// TIA Portal V20 export
// export: Created 2026-10-20T18:56:01.9058217Z, ExportSetting None, DisplayName Totally Integrated Automation Portal, DisplayVersion V20 Update 6, DisplayName TIA Portal Openness, DisplayVersion V20 Update 6, DisplayName TIA Portal Version Control Interface, DisplayVersion V20 Update 6, DisplayName SINAMICS Startdrive Advanced, DisplayVersion V20 SP1, DisplayName SINAMICS Startdrive G130, G150, S120, S150, SINAMICS MV, G220, S200, S210, DisplayVersion V20 SP1, DisplayName SINAMICS Startdrive G110M, G120, G120C, G120D, G120P, G115D, DisplayVersion V20 SP1, DisplayName STEP 7 Professional, DisplayVersion V20 Update 6, DisplayName STEP 7 Safety, DisplayVersion V20 Update 2, DisplayName WinCC Basic/Comfort/Advanced, DisplayVersion V20 Update 6, DisplayName WinCC Unified, DisplayVersion V20 Update 6
VAR_GLOBAL   // PLC tag table "Lock_11"
   Switches_11 AT %IB1576 : Byte;
   "Solenoid Enable_11" AT %Q1504.0 : Bool;
   "Lock Reset_11" AT %Q1505.0 : Bool;
   Lamps_11 AT %QB1503 : Byte;
   Lock_11_Estop_CH1 AT %I1838.2 : Bool;
   Lock_11_Estop_CH2 AT %I1838.3 : Bool;
   Lock_11_Closed_CH2 AT %I1838.1 : Bool;
   Lock_11_Closed_CH1 AT %I1838.0 : Bool;
   Lock_11_Reset_Input1 AT %Q1839.0 : Bool;
   Lock_11_Reset_Input3 AT %Q1839.2 : Bool;
   Lock_11_Reset_Input4 AT %Q1839.3 : Bool;
   Lock_11_Reset_Input2 AT %Q1839.1 : Bool;
   "Guard Position_11" AT %I1577.0 : Bool;
   "Lock Position_11" AT %I1846.0 : Bool;
END_VAR
